ABB RobotStudio station: Pallet_Project_valla_practica.rspag

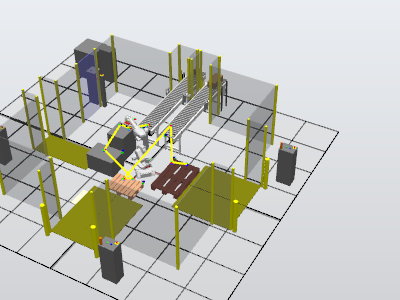
--- station ---
Station Pallet_Project (saved by RobotStudio 24.4.11080.0)
Controller Controler
  mechanical unit ROB_1: IRB1600_10_145__02, 6 joints, base frame (0, 0, 0) mm, rotated rx 0 ry 0 rz 135 deg
Layout (positions relative to the parent item):
  - IRB1600_10_145__02 [mechanism, from %ABB.RobotStudio.Models.IRB1600%\IRB1600_10_145_G_02.rslib] at (0, 0, 0) mm, rotated rx 0 ry 0 rz 135 deg; joint values [0.3434, -0.1552, -0.118, 0, 1.844, -0.442] (rad or m)
  - Half EPAL [part] at (-400, -600, 0) mm, rotated rx 0 ry 0 rz -90 deg, size 600 x 800 x 144 mm
  - ConveyorBox1 [part, from %ABB.RobotStudio.Models.Conveyors%\Conveyor Guide 400.rslib] at (150, 3660, 0) mm, rotated rx 0 ry 0 rz -90 deg
  - ConveyorBox2 [part, from %ABB.RobotStudio.Models.Conveyors%\Conveyor Guide 400.rslib] at (-550, 3660, 0) mm, rotated rx 0 ry 0 rz -90 deg
  - PalletizingVacuumTool [mechanism] at (-560, 265, 1275) mm, rotated rx 180 ry 0 rz 0 deg
      TCP toolVacuum at (0, 0, 175) mm
      links: PalletizingVacuumTool
  - Box1 [part] at (338.5, 3410, 868) mm, size 249 x 499 x 200 mm
  - Box2 [part] at (-353.5, 3575, 868) mm, size 129 x 129 x 200 mm
  - EuroPallet [part, from Components\EuroPalletWood.rslib] at (1400, -600, 0) mm, rotated rx 0 ry 0 rz 90 deg
  - StackingTable [part], size 500 x 600 x 770 mm
  - LinerStand [part], size 800 x 540 x 500 mm
  - SC_Conveyor1 [smart component]
      signals: DO BoxArrived, DI EuroPalletReplaced, DO EuroPalletReplacedOut, DI EuroPalletFull
      connections:
        Source.Executed -> Queue.Enqueue
        PlaneSensor.SensorOut -> Queue.Dequeue
        PlaneSensor.SensorOut -> SC_Conveyor1.BoxArrived
        PlaneSensor.SensorOut -> LogicGate_2.InputA
        LogicGate_2.Output -> Queue_EuroPallet.Enqueue
        LogicGate_2.Output -> Source.Execute
        SimulationEvents.SimulationStarted -> Source.Execute
        SC_Conveyor1.EuroPalletReplaced -> LogicGate_4.InputA
        SC_Conveyor1.EuroPalletFull -> LogicGate_4.InputB
        LogicGate_4.Output -> Queue_EuroPallet.DeleteAll
        LogicGate_4.Output -> SC_Conveyor1.EuroPalletReplacedOut
        Source.Copy => Queue.Back
        Source.Copy => Queue_EuroPallet.Back
    - Source [smart component, from Components\Source.rslib]
        properties: Source=Box1; Copy=(none); Parent=(none); Position=[0.3385 3.39 0.868]; Orientation=[0 0 0]; Transient=true; PhysicsBehavior=-1
    - Queue [smart component, from Components\Queue.rslib]
        properties: Back=(none); Front=(none); Queue={e44fd220-027a-471e-9bb3-a121b85bf4f4};{ee89139f-02ff-44ed-9ba1-277313a75013};{18dc721d-160d-4138-ae65-9469c6fd54a3};{8a7c9217-9ec1-4f6b-adb2-90e3a400ce08};{00ac1772-6055-444c-babb-fd014df5a64d};{22d9b99e-02f4-42e2-875d-e7a2e7a407a6};{801c1d70-c872-49cf-9333-ae7f090aa808};{70a3d2ac-7d8e-4e25-ad4d-efa1d0715e14};{3d190289-ddf5-4821-aefa-1399e7a245df};{fd209546-ad15-4917-a822-45590f893235};{336d7e34-4da5-4704-8767-4e7065a2785d};{a26fb9d1-bd3f-44a5-b61e-f217acd5645d};{35f192af-f0b1-4fcb-92d4-6c5266967521};{7901bdf8-4259-4a58-9fb5-5cf3c990d920};{342c242d-4c7b-4a99-80ec-4606a83008e6};{ba259da1-5c68-49c6-a6dd-ca9a29fb7a6a}; NumberOfObjects=0
    - LinearMover [smart component, from Components\LinearMover.rslib]
        properties: Object=Queue; Direction=[0 -0.001 0]; Speed=0.25; Reference=Global; ReferenceObject=(none)
    - PlaneSensor [smart component, from Components\PlaneSensor.rslib]
        properties: Origin=[0.1885 0.675 0.788]; Axis1=[0.3 0 0]; Axis2=[0 0 0.01]; Tag=(none); SenseMultiple=false; SensedPart=(none)
      - _sensorPart_ [part], size 300 x 0 x 10 mm
    - LogicGate_2 [smart component, from Components\LogicGate.rslib]
        properties: Operator=NOT; Delay=0
    - SimulationEvents [smart component, from Components\SimulationEvents.rslib]
    - Queue_EuroPallet [smart component, from Components\Queue.rslib]
        properties: Back=(none); Front=(none); Queue={ad2057dc-9812-4e01-8eaf-a9764e1c94d2};{23c6148b-879e-4f76-bca6-d4d483c6d4cf};{54fab71e-bcc4-4cca-934a-bbba160b39cc};{b0578ce1-49ea-4c32-a7ca-1e85ec604af9};{947d5054-25d5-43c7-944a-6033d179de93};{94505b46-0998-4fbc-8e5e-e62bbe244ad7};{f8f4ee6a-1769-49de-aeb3-fda26ec8c2f8};{b15d2938-3ac6-4e58-8ecd-de010d23430d};{1b2107f9-d4c6-43db-8eaa-2f076badebbf};{8fdf9589-2ad3-4260-9f23-49ca6aa9f936};{e6f3ceb5-7ecf-422f-9b07-fa91f87616c7};{f8c0f3b0-c392-4387-85be-b0b3c79b7ed2};{b39ef0a3-239a-4eec-87db-20edab27732a};{5504cbc0-0a84-43c9-a60a-8c085a41512d};{4d3e807d-0d48-4360-91da-1f89d28d46d8};{a29bebad-6711-442d-b78a-1822bba72e52};{67d8694a-6ead-419a-ae85-289693a6d2b4};{fe453467-8abc-48a3-b851-8c12c1d7de9d};{6a3e15a0-208f-443f-b6ba-a36fe2c16062};{20e970d1-663c-443e-a64d-d4e9619459f6};{5c8b92e3-60f3-4981-96e7-ca10cb27a842};{db639feb-fd6e-461a-932d-f627d06db2d4};{94b1b66a-00eb-48e1-8857-3db09adf90dc};{618ef0e4-4d6b-4c69-b61e-0bdaa313040e};{043080b5-4091-48b4-bcaf-45ad99666a15};{29caf58f-62f3-4756-8934-f4cc9122e7eb};{7885f061-03ec-4f1c-9005-bd87fa17bd26};{e44fd220-027a-471e-9bb3-a121b85bf4f4};{ee89139f-02ff-44ed-9ba1-277313a75013};{8a7c9217-9ec1-4f6b-adb2-90e3a400ce08};{00ac1772-6055-444c-babb-fd014df5a64d};{22d9b99e-02f4-42e2-875d-e7a2e7a407a6};{801c1d70-c872-49cf-9333-ae7f090aa808};{70a3d2ac-7d8e-4e25-ad4d-efa1d0715e14};{3d190289-ddf5-4821-aefa-1399e7a245df};{fd209546-ad15-4917-a822-45590f893235};{336d7e34-4da5-4704-8767-4e7065a2785d};{a26fb9d1-bd3f-44a5-b61e-f217acd5645d};{35f192af-f0b1-4fcb-92d4-6c5266967521};{7901bdf8-4259-4a58-9fb5-5cf3c990d920};{342c242d-4c7b-4a99-80ec-4606a83008e6}; NumberOfObjects=12
    - LogicGate_4 [smart component, from Components\LogicGate.rslib]
        properties: Operator=AND; Delay=0
  - SC_Gripper [smart component]
      signals: DI Grip
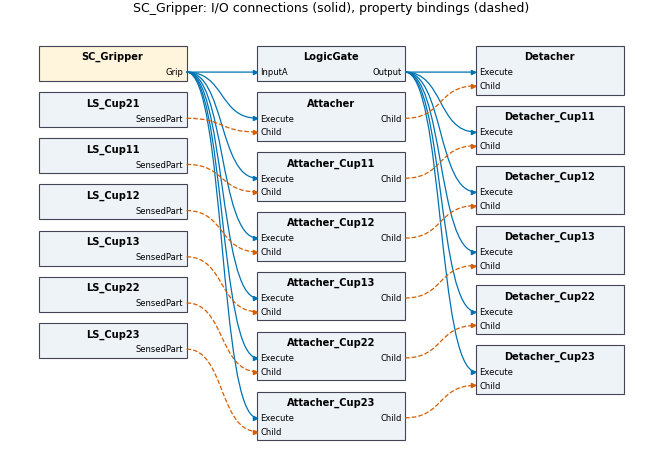
      connections:
        SC_Gripper.Grip -> Attacher.Execute
        SC_Gripper.Grip -> LogicGate.InputA
        LogicGate.Output -> Detacher.Execute
        SC_Gripper.Grip -> Attacher_Cup11.Execute
        LogicGate.Output -> Detacher_Cup11.Execute
        SC_Gripper.Grip -> Attacher_Cup12.Execute
        LogicGate.Output -> Detacher_Cup12.Execute
        SC_Gripper.Grip -> Attacher_Cup13.Execute
        LogicGate.Output -> Detacher_Cup13.Execute
        SC_Gripper.Grip -> Attacher_Cup22.Execute
        LogicGate.Output -> Detacher_Cup22.Execute
        SC_Gripper.Grip -> Attacher_Cup23.Execute
        LogicGate.Output -> Detacher_Cup23.Execute
        LS_Cup21.SensedPart => Attacher.Child
        Attacher.Child => Detacher.Child
        LS_Cup11.SensedPart => Attacher_Cup11.Child
        Attacher_Cup11.Child => Detacher_Cup11.Child
        LS_Cup12.SensedPart => Attacher_Cup12.Child
        Attacher_Cup12.Child => Detacher_Cup12.Child
        LS_Cup13.SensedPart => Attacher_Cup13.Child
        Attacher_Cup13.Child => Detacher_Cup13.Child
        LS_Cup22.SensedPart => Attacher_Cup22.Child
        Attacher_Cup22.Child => Detacher_Cup22.Child
        LS_Cup23.SensedPart => Attacher_Cup23.Child
        Attacher_Cup23.Child => Detacher_Cup23.Child
    - LS_Cup21 [smart component, from Components\LineSensor.rslib] at (190, 265, 153.5) mm, rotated rx 0 ry 0 rz 45 deg
        properties: Start=[-0.597509982704304 0.689429996191639 0.956499992313755]; End=[-0.597509981617333 0.689429995104668 0.924499992313755]; Length=0.032; Radius=0.00331491712707182; Tag=(none); SenseMultiple=false; SensedPart=(none); SensedPoint=[0 0 0]
      - _sensorPart_ [part], size 6.4 x 6.4 x 32 mm
    - Attacher [smart component, from Components\Attacher.rslib]
        properties: Parent=PalletizingVacuumTool; Flange=0; Child=(none); Mount=false; Offset=[0 0 0]; Orientation=[0 0 0]
    - Detacher [smart component, from Components\Detacher.rslib]
        properties: Child=(none); KeepPosition=true
    - LogicGate [smart component, from Components\LogicGate.rslib]
        properties: Operator=NOT; Delay=0
    - LS_Cup11 [smart component, from Components\LineSensor.rslib] at (190, 265, 153.5) mm, rotated rx 0 ry 0 rz 45 deg
        properties: Start=[-0.68943 0.59751 0.9565]; End=[-0.68943 0.59751 0.9245]; Length=0.032; Radius=0.00331; Tag=(none); SenseMultiple=false; SensedPart=(none); SensedPoint=[0 0 0]
      - _sensorPart_ [part], size 6.6 x 6.6 x 32 mm
    - LS_Cup12 [smart component, from Components\LineSensor.rslib] at (190, 265, 153.5) mm, rotated rx 0 ry 0 rz 45 deg
        properties: Start=[-0.57629 0.48437 0.9565]; End=[-0.57629 0.48437 0.9245]; Length=0.032; Radius=0.00331; Tag=(none); SenseMultiple=false; SensedPart=(none); SensedPoint=[0 0 0]
      - _sensorPart_ [part], size 6.6 x 6.6 x 32 mm
    - LS_Cup13 [smart component, from Components\LineSensor.rslib] at (190, 265, 153.5) mm, rotated rx 0 ry 0 rz 45 deg
        properties: Start=[-0.46315 0.37123 0.9565]; End=[-0.46315 0.37123 0.9245]; Length=0.032; Radius=0.00331; Tag=(none); SenseMultiple=false; SensedPart=(none); SensedPoint=[0 0 0]
      - _sensorPart_ [part], size 6.6 x 6.6 x 32 mm
    - LS_Cup22 [smart component, from Components\LineSensor.rslib] at (190, 265, 153.5) mm, rotated rx 0 ry 0 rz 45 deg
        properties: Start=[-0.48437 0.57629 0.9565]; End=[-0.48437 0.57629 0.9245]; Length=0.032; Radius=0.00331; Tag=(none); SenseMultiple=false; SensedPart=(none); SensedPoint=[0 0 0]
      - _sensorPart_ [part], size 6.6 x 6.6 x 32 mm
    - LS_Cup23 [smart component, from Components\LineSensor.rslib] at (190, 265, 153.5) mm, rotated rx 0 ry 0 rz 45 deg
        properties: Start=[-0.37123 0.46315 0.9565]; End=[-0.37123 0.46315 0.9245]; Length=0.032; Radius=0.00331; Tag=(none); SenseMultiple=false; SensedPart=(none); SensedPoint=[0 0 0]
      - _sensorPart_ [part], size 6.6 x 6.6 x 32 mm
    - Attacher_Cup11 [smart component, from Components\Attacher.rslib]
        properties: Parent=PalletizingVacuumTool; Flange=0; Child=(none); Mount=false; Offset=[0 0 0]; Orientation=[0 0 0]
    - Detacher_Cup11 [smart component, from Components\Detacher.rslib]
        properties: Child=(none); KeepPosition=true
    - Attacher_Cup12 [smart component, from Components\Attacher.rslib]
        properties: Parent=PalletizingVacuumTool; Flange=0; Child=(none); Mount=false; Offset=[0 0 0]; Orientation=[0 0 0]
    - Detacher_Cup12 [smart component, from Components\Detacher.rslib]
        properties: Child=(none); KeepPosition=true
    - Attacher_Cup13 [smart component, from Components\Attacher.rslib]
        properties: Parent=PalletizingVacuumTool; Flange=0; Child=(none); Mount=false; Offset=[0 0 0]; Orientation=[0 0 0]
    - Detacher_Cup13 [smart component, from Components\Detacher.rslib]
        properties: Child=(none); KeepPosition=true
    - Attacher_Cup22 [smart component, from Components\Attacher.rslib]
        properties: Parent=PalletizingVacuumTool; Flange=0; Child=(none); Mount=false; Offset=[0 0 0]; Orientation=[0 0 0]
    - Detacher_Cup22 [smart component, from Components\Detacher.rslib]
        properties: Child=(none); KeepPosition=true
    - Attacher_Cup23 [smart component, from Components\Attacher.rslib]
        properties: Parent=PalletizingVacuumTool; Flange=0; Child=(none); Mount=false; Offset=[0 0 0]; Orientation=[0 0 0]
    - Detacher_Cup23 [smart component, from Components\Detacher.rslib]
        properties: Child=(none); KeepPosition=true
  - SC_Conveyor2 [smart component]
      signals: DO BoxArrived, DI HalfPalletReplaced, DI HalfPalletFull, DO HalfPalletReplacedOut
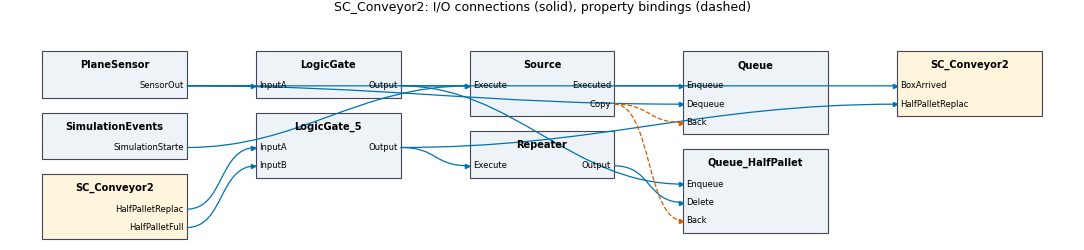
      connections:
        Source.Executed -> Queue.Enqueue
        PlaneSensor.SensorOut -> Queue.Dequeue
        PlaneSensor.SensorOut -> SC_Conveyor2.BoxArrived
        PlaneSensor.SensorOut -> LogicGate.InputA
        SimulationEvents.SimulationStarted -> Source.Execute
        LogicGate.Output -> Queue_HalfPallet.Enqueue
        LogicGate.Output -> Source.Execute
        Repeater.Output -> Queue_HalfPallet.Delete
        SC_Conveyor2.HalfPalletReplaced -> LogicGate_5.InputA
        SC_Conveyor2.HalfPalletFull -> LogicGate_5.InputB
        LogicGate_5.Output -> Repeater.Execute
        LogicGate_5.Output -> SC_Conveyor2.HalfPalletReplacedOut
        Source.Copy => Queue.Back
        Source.Copy => Queue_HalfPallet.Back
    - Source [smart component, from Components\Source.rslib]
        properties: Source=Box2; Copy=(none); Parent=(none); Position=[-0.3535 3.575 0.868]; Orientation=[0 0 0]; Transient=true; PhysicsBehavior=-1
    - Queue [smart component, from Components\Queue.rslib]
        properties: Back=(none); Front=(none); Queue={d41f34b8-4a20-475c-95ba-460bc2504caf};{5a16ad96-9ff6-44fe-ab59-6bd35466d4d1};{0f18d6dc-c4e6-4c44-9757-559d16fce4ae};{b2c7b4bf-0d60-42df-8ee4-abc0a1068e12};{8d30a67c-a063-4d22-a747-3e9a99cdef41};{1409c1e2-dbf3-49bd-b776-9bd8588f9165};{e3acce53-8455-4384-b1ac-df89878ccd5c};{87db3190-4758-4831-8d2c-d9fdcd68b36e};{469258bd-729a-49fe-bc80-31f695b1b400};{4c1b5bae-9eaf-40c3-874b-2538b6841d7a};{46ba244e-445c-470d-b6ca-5e376dcf2b7e};{e5ec3e26-f6d7-4e6f-b347-541b5d6ec99e}; NumberOfObjects=0
    - LinearMover [smart component, from Components\LinearMover.rslib]
        properties: Object=Queue; Direction=[0 -0.001 0]; Speed=0.25; Reference=Global; ReferenceObject=(none)
    - PlaneSensor [smart component, from Components\PlaneSensor.rslib]
        properties: Origin=[-0.5035 0.675 0.788]; Axis1=[0.3 0 0]; Axis2=[0 0 0.01]; Tag=(none); SenseMultiple=false; SensedPart=(none)
      - _sensorPart_ [part], size 300 x 0 x 10 mm
    - LogicGate [smart component, from Components\LogicGate.rslib]
        properties: Operator=NOT; Delay=0
    - SimulationEvents [smart component, from Components\SimulationEvents.rslib]
    - Queue_HalfPallet [smart component, from Components\Queue.rslib]
        properties: Back=(none); Front=(none); Queue={f5edb1ce-3bf5-426a-a389-0b0047efa949};{5ce0816a-b692-43c6-82f7-492eb3fc1c7c};{ad3ef4b5-2c59-4daa-9658-0c77e5efb67d};{c9c476d0-74ff-4b18-bfb3-2d6c852b8493};{1bf865c6-1649-4319-b5ff-cd81faaa6069};{f626778c-15a6-4059-b27a-7c8f9da4f34f};{a60dd0dd-490e-48fe-bb32-16f415136b44};{4ec9b3b2-e4a8-4d14-aea0-9552a35d2afd};{38bc6a68-8d9e-44a7-a5f0-badb214ea710};{f9543542-377a-43f1-9613-018dced76680};{486b4c2f-b225-4486-b430-5ab7d813c599};{7da52d9e-9053-4b1a-839c-0aedc5495cc7};{c2400356-fde5-4523-9dc7-d26788098951};{75099568-1fe6-4c34-8328-63fd42144c3b};{8ca6c374-2d39-4938-8324-38c48ae4f51d};{f3c160ab-6f5f-460b-8b54-c2c3b0bc175f};{1c289510-9a29-4e1c-b603-54b7a0027260};{d39da69b-e59a-4ace-85a5-bba54583b01c};{bc328c62-4bf3-4a57-965c-0c93e0ee296d};{60f4dcb3-d366-4d0b-b05a-5b2073fcd9e8};{44334a49-cf52-4d95-9964-3bb568ce732d};{f9240695-1965-47e5-bcd4-644ec5904899};{72a970fd-f238-4ac5-b811-00686975bc20};{bd297b2a-4ad7-44fa-87c8-1ac40b0d2fbf};{3dafa88d-62b0-429f-9c75-c8c7bde09fc6};{a7d8f176-4e9d-4819-8805-982bee0c310d};{72ae6bb6-3373-4f60-a321-dfdc0981c562};{fff16105-3d56-4b21-a888-399904fd95d4};{56e4abf9-acd4-4a00-b067-52a58200d221};{2eb8ae55-b553-4f83-b65d-07c27c701dd6};{dfb05241-1220-45e8-b584-1559777c0125};{49a2c23a-27ea-4b0b-af5c-f9d01014f642};{0adfb5d7-4fd0-41be-8361-c42c9d28ca51};{8cf74624-f46b-49ca-a524-038ddb88ba0f};{bde2cdc4-b3e4-48fe-8333-d64185b5a8e7};{d17564c2-89d4-4b4f-8596-5dca9165a286};{6fec26e7-cb1b-4d74-b4a6-8ed7a2eb81a6};{e04d8697-cc19-4df5-b7fa-dff41516820c};{134714af-70a5-49a3-8b99-ea847d1ef329};{23aa8eff-aaeb-4079-b6e6-9fe5f0b7799c};{0091a76d-e23e-4382-9bf3-a427b049953f};{fdc2abc9-40b2-462e-8472-b1d156765a68};{8dc86a38-8dcf-454b-a79a-3f5e6d46a581};{f9226736-fe9f-4ce5-82b5-97fc8f487c87};{8d0584df-2d5d-4d5a-bd5b-c865cb85c145};{fef2818e-b6b9-47fe-bf8a-83543bb000b1};{5ac98beb-c6da-4ea7-80b2-93f7dacce3e5};{443aad51-6408-442e-915b-2ecfdc577e14};{51b93794-f199-43f0-a14e-6aec3c171668};{885be8a6-b854-423c-907a-f456456dba07};{dcbbb2a9-79f1-4094-9b60-3ac8a0070454};{86281ae9-2d9e-4987-a35e-6d6a445e8875};{9f234810-50d8-438d-8980-298a5844ac16};{4c457525-5ea0-4a08-bfa0-e2a51e8a57a9};{d60c358c-9baa-495a-a755-dc91e6e5630d};{cba8d61a-9576-424b-b333-8920ed1679e6};{fffcb6aa-6454-497e-a713-529b874f7300};{8c292b69-8603-4861-ab75-8c5041fc1228};{be74d22e-2a24-4d51-b9be-30cb4581f5e4};{9c8c849d-9d7a-4314-9edc-0c9679818308};{51cbe104-3a08-4083-a326-34fc650c90a2};{8d9adc3a-e0d0-484f-8727-84b992719000};{9a2b47ee-5540-43de-9a30-89f96a258b35};{cfb929ec-bf51-45d3-8071-aea9b14bf075};{867175b9-70b9-45ce-970c-131187ba34ca};{173082af-f5ae-4239-8a69-7ad684951e00};{b2c9da23-dceb-4407-8f95-0d503246dac3};{f0464754-db31-42ef-9c41-8ce46a4a0971};{6b29df5c-760d-4911-84dd-92d25b30bb71};{8cf0ae3d-fbb1-4655-8db9-abf8850d857b};{fcdbf145-8b27-4e5e-9241-3719648eab1d};{78faf9d5-81df-4a41-87f3-b1a514ef17c7};{3a4d91ff-54a0-485c-9c99-c5554510e37a};{c01a110e-561d-45dd-b1c3-10d79a4111a8};{63ad2c6d-e580-44e3-9dfc-7106564b7944};{ccc00ef2-4c06-4459-824e-6f17fc3bacb7};{b81e233c-b00c-4cd7-b93a-2cecac8f8dc1};{398e0c88-f727-4b42-8f39-aaa6835500b7};{fc631786-067a-487d-abac-51fcb0c6dd41};{cf6ca633-09f3-4f3b-9435-b43791280bff};{74bed72d-6a54-4305-87bd-9ad3015ece89};{bb2cc45e-a4eb-4ab2-9ef7-f371e7fbe706};{dd82f376-2e09-4208-84ad-5816bed92574};{e392904e-f13d-4939-a056-7304ff0c878c};{3e44c1eb-892b-48b7-9eef-a2eb6a338ec4};{67a95a53-b6c9-4e7f-9fd4-7782a33b0ce9};{b907a4a1-1349-44c4-99ca-3ea2b14844a2};{27bb147c-485e-4ba4-8918-f2e2468aa20b};{4158548c-0e01-4059-887d-ce75515d9624};{bdcc830f-a4a4-4608-9c6a-3968c3b56955};{8ac99da1-daa1-4239-8c24-2cbcd0fbbccf};{eceb8029-a656-40f5-a7a3-28283ded6e47};{06ec9c8e-bd56-4499-906c-965bdc743b38};{bc8629f4-be69-483d-a42b-bd5694970e3a};{91c33ad6-79d6-4ff7-b807-aaf3d283071a};{bbff1efe-9f6d-4f6e-9e11-7159709d58b9};{d8345c1f-8548-4957-9dd2-2c7a65aadcb5};{297050bf-6bdd-4149-9774-639d35df4273};{9047bf3c-f537-46c2-88b1-9fd2d5954a0b};{5951cc55-a535-4f63-8005-57734053514f};{4bb3aaf8-1744-440d-8239-fce36f67cc2c};{eb7c6c5d-8b86-4d0e-b965-01e8cc90c395};{da949c7c-7130-455a-a5de-886672c52ec3};{04b934b1-2ca6-4947-808f-8dc968a55eb4};{d4940027-1ade-4406-ae0f-2cc92eccc776};{37dc3e2f-17e0-406e-80b6-d473aa1734f3};{09cf0d3f-945d-4baa-a296-e9bd267df3af};{8a94d3e3-b0e3-42c4-90bd-ba639180af74};{049eaf7e-723f-484a-b080-48153e5693e0};{2c2227db-366e-4824-818a-8891fec9d39b};{78a4912a-e493-4427-95eb-ed4a7e141f53};{8b1769a4-052b-4f7f-be48-9c2315e00515};{4bb9eccd-54a8-444b-8b85-f69dc35199f7};{5d771788-ec0f-48bc-9cbe-993fb932c8ea};{021fadd8-996c-49c9-9ff6-8a460f8c358b};{e61d541c-af94-4f27-b95d-aac3b95a1cd9};{a0819d77-e800-4559-87f4-c656405fa595};{003f191f-efb3-43bb-b7aa-33133ee6defd};{3abac3eb-5c5c-4177-b0e4-5f71daa2fcd7};{f4938c82-19bc-4592-9d12-63feb2c87ac4};{2b776e4a-67ea-499c-995e-bce8af0160a7};{c9a77fd9-e2d1-4dbf-8d0e-8377c4665448};{62bb8355-d295-4471-b563-b6f46f05c8b1};{55201944-7d05-43e8-bd24-433bd506e7b6};{76821f68-2096-4060-b9d6-b9517b2f6dc5};{e09ad2c9-6668-417d-a6ce-db14256207b6};{ca102da5-219d-413a-ab81-6e9821c26e06};{c588302c-8cce-44a8-91f3-143c0654eb27};{2202393d-e22d-4f8c-8a1d-1cc72ba5cca5};{be80ae30-a6c8-4766-bc6b-bfe80846e161};{25475f3f-ef68-45ff-aa3c-0ea04c10e4e7};{498aca50-8032-4c24-8147-7ec56c07f7a0};{b4a07b3f-831d-4f53-9343-c16642fe3bc1};{8bd52ab4-c09d-4b2d-8603-56cbb3c77529};{6f1069cf-970f-4855-ba49-8ae785987118};{b667b62f-e5f1-478a-9bad-dc3725da1d04};{86e8e265-466a-4a6e-8b5e-b128819dda1c};{4df69d20-688f-43ef-bee0-112974bed187};{182f9b53-f0c9-4414-a7de-97eac4ce486a};{514b0f5e-2197-4430-9c07-cfb19e0d92ad};{359ebd0e-6711-4070-a5d3-939e22007801};{d67847b8-c0ad-4246-ba67-b0d24865206c};{197fb8bb-a523-4e0e-8be7-47cc1723a988};{142dd6b6-47a3-4a32-99f8-9706d11eb229};{1a8963b6-e72b-4e55-95a7-15d5212af876};{42897a06-6f96-425a-a387-4cefe2eac35b};{d78e4ef6-3fce-473d-bfe7-e529abd3d695};{e0b062dd-5846-40f4-b32c-2a1ab6da1894};{4c4aa1cf-e61f-45c1-9c13-55311062428a};{a0d6a9a4-70e0-4c3a-ae7d-eaf5e5bb2112};{bc16083c-a858-482a-a879-7c8861b2473f};{64ab26ad-0b46-4ced-ab7f-1cfee37682ad};{2165d0dd-c254-4ebf-83cc-be68d523d748};{44491ebe-5cdd-46fe-a821-5ec7c79b16a0};{ddfa3b39-85f7-4855-9203-7f7a6cdd8093};{137fe74d-152f-4b74-9f93-d403c4354bb3};{82ca252e-23ba-4001-8e89-7b23c4c78f2e};{062cf830-d27c-401d-a518-3a9fb83d9537};{610befe8-cd72-44d2-af6b-444eaea3df38};{cf0b5eb3-bda2-46b1-b486-9a887917bee5};{a53ebe9a-d0a3-4afd-b901-97852e5709fd};{8b5126a5-3700-41cc-bd9b-a335d093d62b};{1a031046-3bf3-47b0-bf1d-63f834d0f0bf};{32ae9498-3575-4e70-954e-9800b2c7ed18};{ee3cbed5-90f6-47a6-8d41-8a31a6a9b52f};{f52f3a91-5bd6-47b6-a1f8-92ea9cad0f19};{b2f50ce9-01bf-4326-9e7f-81a685c29d51};{db908664-ce90-4d8d-99e6-8cad1d25b072};{ce174d6d-3e8c-4abc-807c-2e034a05442b};{6b3f855e-a78e-40d1-a8e8-dc264647088d};{cde41289-1748-48b7-acac-ba93367ef0bd};{23d0bcac-3df5-4d02-9989-7a0bd57a2c5a};{7d6ef79f-31a3-4faa-a3c8-24190ad66021};{148a4a69-c3f4-4709-9c4e-248710d37209};{3a43107f-6ec5-42b1-bdab-65f53844f08b};{688ca237-9237-4c0d-9f6a-943bdaf2a54e};{b0c649b2-1e95-4926-b3f4-7de3359bf184};{775c86bc-3b84-4fb2-a4b9-0c2b4654e980};{d13aeccf-57c6-48c5-8ccb-e0d83af0bf52};{b23f60bf-e49d-4af6-aa11-454509134c6f};{0a5e5d93-42f5-44d1-80bb-87a9dcd65f82};{03917fb8-4550-48ea-aade-cad2296182d4};{69fc404e-23e5-4586-8106-722a8d502888};{efd93624-9dc8-470c-9ca5-761da3b13f64};{3161c526-c456-4198-a8e9-6ba9dc97d08d};{1f8ccdfc-77be-4eb2-b50b-b6f397d92aac};{cb468d26-4eaa-493f-84ab-65bfcf757383};{bd96b98c-b60d-47b5-9e29-6a1dfadd5ba3};{35cfaa90-f083-49e1-b726-d654efc82f59};{60633137-d3a6-410f-a68f-c3960af01eec};{b8faed0a-d8df-4dd7-a7c6-c20d690a082c};{469fa596-a3ad-4a84-8b8e-6f04cb45c4e6};{543f5b18-19fb-410f-92c3-c1199be26dff};{1f728d5f-b843-4df0-b352-629d14987f1c};{12323632-ef84-4060-aa52-b2f1987c73f3};{062735fc-4a51-4d85-95c2-a683477f8e45};{444b3eac-f57f-4356-8db0-63ce6624c93d};{325a86c2-b1da-40af-a81a-eb00a2886e08};{73c79afd-8798-467b-80dd-9e32e888d88c};{f243e6a9-0264-46d4-8a6c-a8c2b4c42193};{f7d0602e-30eb-44b6-b654-6cdc5756be59};{ad2ed4ca-30e0-4614-a0d8-f4fea7ef6fce};{bab6a964-a4d0-4eed-9c33-fa686721e8e3};{fb67aacc-6733-43ed-a4db-7a6425d2d60c};{6421a31f-3a82-4b20-9081-df48bb7907b5};{8ff8c115-8e7b-4406-a53a-edf3873335b8};{5ac3eee3-ab48-4a86-8294-3ac57f94e03f};{d41f34b8-4a20-475c-95ba-460bc2504caf};{5a16ad96-9ff6-44fe-ab59-6bd35466d4d1};{0f18d6dc-c4e6-4c44-9757-559d16fce4ae};{b2c7b4bf-0d60-42df-8ee4-abc0a1068e12};{8d30a67c-a063-4d22-a747-3e9a99cdef41};{1409c1e2-dbf3-49bd-b776-9bd8588f9165};{e3acce53-8455-4384-b1ac-df89878ccd5c};{87db3190-4758-4831-8d2c-d9fdcd68b36e};{469258bd-729a-49fe-bc80-31f695b1b400};{4c1b5bae-9eaf-40c3-874b-2538b6841d7a};{46ba244e-445c-470d-b6ca-5e376dcf2b7e}; NumberOfObjects=78
    - Repeater [smart component, from Components\Repeater.rslib]
        properties: Count=72
    - LogicGate_5 [smart component, from Components\LogicGate.rslib]
        properties: Operator=AND; Delay=0
  - Liner_01 [part] at (-900, -2000, 0) mm, size 800 x 540 x 10 mm
  - SC_Liners [smart component]
      signals: DI LinersRefilled, DI LinerStackEmpty, DI PalletReplaced, DO LinersRefilledOut
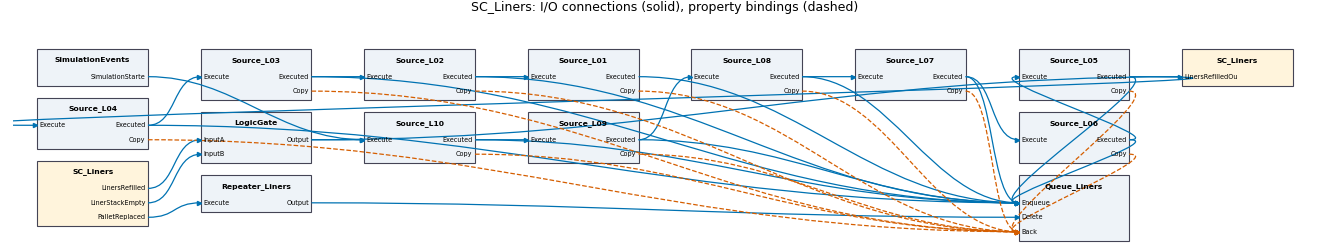
      connections:
        SimulationEvents.SimulationStarted -> Source_L10.Execute
        Source_L10.Executed -> Queue_Liners.Enqueue
        Source_L10.Executed -> Source_L09.Execute
        Source_L09.Executed -> Queue_Liners.Enqueue
        Source_L09.Executed -> Source_L08.Execute
        Source_L08.Executed -> Queue_Liners.Enqueue
        Source_L08.Executed -> Source_L07.Execute
        Source_L07.Executed -> Queue_Liners.Enqueue
        Source_L07.Executed -> Source_L06.Execute
        Source_L06.Executed -> Queue_Liners.Enqueue
        Source_L06.Executed -> Source_L05.Execute
        Source_L05.Executed -> Queue_Liners.Enqueue
        Source_L05.Executed -> Source_L04.Execute
        Source_L04.Executed -> Queue_Liners.Enqueue
        Source_L04.Executed -> Source_L03.Execute
        Source_L03.Executed -> Queue_Liners.Enqueue
        Source_L03.Executed -> Source_L02.Execute
        Source_L02.Executed -> Queue_Liners.Enqueue
        Source_L02.Executed -> Source_L01.Execute
        Source_L01.Executed -> Queue_Liners.Enqueue
        SC_Liners.LinersRefilled -> LogicGate.InputA
        SC_Liners.LinerStackEmpty -> LogicGate.InputB
        LogicGate.Output -> SC_Liners.LinersRefilledOut
        LogicGate.Output -> Source_L10.Execute
        SC_Liners.PalletReplaced -> Repeater_Liners.Execute
        Repeater_Liners.Output -> Queue_Liners.Delete
        Source_L10.Copy => Queue_Liners.Back
        Source_L09.Copy => Queue_Liners.Back
        Source_L08.Copy => Queue_Liners.Back
        Source_L07.Copy => Queue_Liners.Back
        Source_L06.Copy => Queue_Liners.Back
        Source_L05.Copy => Queue_Liners.Back
        Source_L04.Copy => Queue_Liners.Back
        Source_L03.Copy => Queue_Liners.Back
        Source_L02.Copy => Queue_Liners.Back
        Source_L01.Copy => Queue_Liners.Back
    - Source_L10 [smart component, from Components\Source.rslib]
        properties: Source=Liner_01; Copy=(none); Parent=(none); Position=[-1.3 -0.7 0.59]; Orientation=[0 0 0]; Transient=true; PhysicsBehavior=-1
    - Source_L09 [smart component, from Components\Source.rslib]
        properties: Source=Liner_01; Copy=(none); Parent=(none); Position=[-1.3 -0.7 0.58]; Orientation=[0 0 0]; Transient=true; PhysicsBehavior=-1
    - Queue_Liners [smart component, from Components\Queue.rslib]
        properties: Back=(none); Front=(none); Queue={4b76874b-49d8-40e7-b1bf-01d8cc753daf};{f1bc3993-1843-4745-a916-cd233907ef8f};{7d1f5471-804d-47e8-8c82-babb94078c4f};{35f64396-636a-40cf-85a6-257e77a6ae60};{2aedaf41-8ae8-41b0-9db2-9de3ceaf795b};{436fe240-c7f2-42eb-89c0-1cd4aff7e3ff};{e7949e0b-2972-403e-9743-54dc0693f87f};{59bd0fcf-8828-44fb-b45a-84ebd2dc8c3d};{59a7902e-96f8-4e0e-b708-dc1c92c26f66};{1f249118-cd38-42be-b8a7-d3254198917b};{33f64cea-21b7-4476-9a21-b1850c845c4c};{6d880d10-0093-43e7-8014-139534ada452};{8432c400-4781-49f7-aa39-fa2dc6e98a0f};{61e97684-8218-4ac6-a060-0ca69cab5273};{78371439-59e8-482d-8147-9dece47c4b3d};{5351f5ec-037c-4625-be08-d259f2f0dab9};{1728b901-d880-497f-a9dc-fc428da0f52d};{94273ab4-5060-46c3-80b2-362935833b91};{3e6b5fa6-26e1-42c5-aada-9e85978ab4cf};{89a16311-d9f3-4be9-874c-e3d1f0939d0f};{01a3968c-dc38-41a8-821e-9eb7eb9ddcb6};{f6651478-43f4-42ca-bae1-f1f503b6b42a};{2f17a5c0-632c-4a5a-aea8-f6e212c5841b};{69ef7725-acb4-4562-810a-a97a14cbd53c};{704c2d3b-24d3-475f-8d25-b6b26e7fec9c};{f2ed20fd-a82f-4770-a0af-12c07cfbfa73};{d8dcd6ae-656a-4bcc-8399-251caf5a0e2f};{4f1be6df-21fc-4212-9b62-51a6ddf46789};{f83a54dd-86e1-4b51-ad4c-f3092acc29ee};{534771e2-1ace-4b39-b107-fcece75fcd88};{006ab1e9-1667-49eb-a3fc-9daf3d261695};{5cff699e-b7b2-4f06-b0dd-3aa3a2565d54};{62b4127a-2a9b-4d56-a22d-ac07527ab970};{72a0e263-fa92-4955-bee8-75cd8e7bcda3};{2f5c7ce6-cc96-4025-8b6f-42fc8d1c53de};{a007f585-8c80-40f3-9f22-79fa01fd41be};{7214a086-acb6-4dc9-80a5-5db08c6fb4b9};{12bb64d4-b495-4b48-a9c8-db9791f029e3};{32b5cfa5-8504-4b44-a4bf-b1b8b1e80030};{60a53e66-30e6-4fde-a9d2-765474ab08f2};{31019e2a-21cb-4e2c-9cdb-7de64fe533e9};{09e6c226-ece6-4f81-9df3-2592efd7026c}; NumberOfObjects=10
    - SimulationEvents [smart component, from Components\SimulationEvents.rslib]
    - Source_L08 [smart component, from Components\Source.rslib]
        properties: Source=Liner_01; Copy=(none); Parent=(none); Position=[-1.3 -0.7 0.57]; Orientation=[0 0 0]; Transient=true; PhysicsBehavior=-1
    - Source_L07 [smart component, from Components\Source.rslib]
        properties: Source=Liner_01; Copy=(none); Parent=(none); Position=[-1.3 -0.7 0.56]; Orientation=[0 0 0]; Transient=true; PhysicsBehavior=-1
    - Source_L06 [smart component, from Components\Source.rslib]
        properties: Source=Liner_01; Copy=(none); Parent=(none); Position=[-1.3 -0.7 0.55]; Orientation=[0 0 0]; Transient=true; PhysicsBehavior=-1
    - Source_L05 [smart component, from Components\Source.rslib]
        properties: Source=Liner_01; Copy=(none); Parent=(none); Position=[-1.3 -0.7 0.54]; Orientation=[0 0 0]; Transient=true; PhysicsBehavior=-1
    - Source_L04 [smart component, from Components\Source.rslib]
        properties: Source=Liner_01; Copy=(none); Parent=(none); Position=[-1.3 -0.7 0.53]; Orientation=[0 0 0]; Transient=true; PhysicsBehavior=-1
    - Source_L03 [smart component, from Components\Source.rslib]
        properties: Source=Liner_01; Copy=(none); Parent=(none); Position=[-1.3 -0.7 0.52]; Orientation=[0 0 0]; Transient=true; PhysicsBehavior=-1
    - Source_L02 [smart component, from Components\Source.rslib]
        properties: Source=Liner_01; Copy=(none); Parent=(none); Position=[-1.3 -0.7 0.51]; Orientation=[0 0 0]; Transient=true; PhysicsBehavior=-1
    - Source_L01 [smart component, from Components\Source.rslib]
        properties: Source=Liner_01; Copy=(none); Parent=(none); Position=[-1.3 -0.7 0.5]; Orientation=[0 0 0]; Transient=true; PhysicsBehavior=-1
    - LogicGate [smart component, from Components\LogicGate.rslib]
        properties: Operator=AND; Delay=0
    - Repeater_Liners [smart component, from Components\Repeater.rslib]
        properties: Count=2
  - Door_Maintenance [part], size 20 x 800 x 2000 mm
  - LightCurtain_EuroPallet_Emitter [part], size 50 x 50 x 2000 mm
  - LightCurtain_EuroPallet_Receiver [part], size 50 x 50 x 2000 mm
  - LightCurtain_HalfPallet_Emitter [part], size 50 x 50 x 2000 mm
  - LightCurtain_HalfPallet_Receiver [part], size 50 x 50 x 2000 mm
  - LightCurtain_LinerBay_Emitter [part], size 50 x 50 x 2000 mm
  - LightCurtain_LinerBay_Receiver [part], size 50 x 50 x 2000 mm
  - LightCurtain_Conv1_Emitter [part], size 50 x 50 x 450 mm
  - LightCurtain_Conv1_Receiver [part], size 50 x 50 x 450 mm
  - LightCurtain_Conv2_Emitter [part], size 50 x 50 x 450 mm
  - LightCurtain_Conv2_Receiver [part], size 50 x 50 x 450 mm
  - MutingSensor_Conv1_A [part], size 30 x 30 x 900 mm
  - MutingSensor_Conv1_B [part], size 30 x 30 x 900 mm
  - MutingSensor_Conv2_A [part], size 30 x 30 x 900 mm
  - MutingSensor_Conv2_B [part], size 30 x 30 x 900 mm
  - SafetyMat_EuroPallet [part], size 1650 x 1800 x 15 mm
  - SafetyMat_HalfPallet [part], size 1500 x 1850 x 15 mm
  - SafetyMat_LinerBay [part], size 1750 x 740 x 15 mm
  - PalletStop_Euro_1 [part], size 40 x 100 x 80 mm
  - PalletStop_Euro_2 [part], size 40 x 100 x 80 mm
  - PalletStop_Half_1 [part], size 100 x 40 x 80 mm
  - PalletStop_Half_2 [part], size 100 x 40 x 80 mm
  - OperatorStation_EuroPallet [part], size 400 x 300 x 1100 mm
  - OperatorStation_HalfPallet [part], size 400 x 300 x 1100 mm
  - OperatorStation_LinerBay [part], size 400 x 300 x 1100 mm
  - OperatorStation_General [part], size 400 x 300 x 1100 mm
  - OperatorStation_Door [part], size 300 x 300 x 1100 mm
  - EStopPost_Inside [part], size 100 x 100 x 1100 mm
  - IRC5_Cabinet [part], size 725 x 710 x 970 mm
  - DoorSensor_Eden_Actuator [part], size 30 x 40 x 60 mm
  - DoorSensor_Eden_Sensor [part], size 30 x 40 x 60 mm
  - EStopBase_EuroPallet [part], size 80 x 80 x 5 mm
  - EStopBase_HalfPallet [part], size 80 x 80 x 5 mm
  - EStopBase_LinerBay [part], size 80 x 80 x 5 mm
  - EStopBase_General [part], size 80 x 80 x 5 mm
  - EStopBase_Door [part], size 80 x 80 x 5 mm
  - EStopBase_Inside [part], size 80 x 80 x 5 mm
  - Bumper_EuroPallet_1 [part], size 114 x 114 x 1000 mm
  - Bumper_EuroPallet_2 [part], size 114 x 114 x 1000 mm
  - Bumper_HalfPallet_1 [part], size 114 x 114 x 1000 mm
  - Bumper_HalfPallet_2 [part], size 114 x 114 x 1000 mm
  - MutingLamp_Conv1 [part], size 60 x 60 x 100 mm
  - MutingLamp_Conv2 [part], size 60 x 60 x 100 mm
  - Lamp_EuroPalletFull [part], size 60 x 59.8 x 200 mm
  - Lamp_HalfPalletFull [part], size 60 x 59.8 x 200 mm
  - Lamp_LinerStackEmpty [part], size 60 x 59.8 x 200 mm
  - Button_EuroPalletReplaced [part], size 40 x 39.9 x 20 mm
  - Button_HalfPalletReplaced [part], size 40 x 39.9 x 20 mm
  - Button_LinersRefilled [part], size 40 x 39.9 x 20 mm
  - ResetButton_EuroPallet [part], size 40 x 39.9 x 20 mm
  - ResetButton_HalfPallet [part], size 40 x 39.9 x 20 mm
  - ResetButton_LinerBay [part], size 40 x 39.9 x 20 mm
  - ResetButton_Door [part], size 40 x 39.9 x 20 mm
  - EStop_EuroPallet [part], size 40 x 40 x 30 mm
  - EStop_HalfPallet [part], size 40 x 40 x 30 mm
  - EStop_LinerBay [part], size 40 x 40 x 30 mm
  - EStop_General [part], size 40 x 40 x 30 mm
  - EStop_Door [part], size 40 x 40 x 30 mm
  - EStop_Inside [part], size 40 x 40 x 30 mm
  - Safety_Fence [graphiccomponentgroup]
    - Fence_Corridor_Euro_1 [part], size 500 x 20 x 2000 mm
    - Fence_Corridor_Euro_2 [part], size 500 x 20 x 2000 mm
    - Fence_Corridor_Half_1 [part], size 20 x 500 x 2000 mm
    - Fence_Corridor_Half_2 [part], size 20 x 500 x 2000 mm
    - Fence_Corridor_Liner_1 [part], size 500 x 20 x 2000 mm
    - Fence_Corridor_Liner_2 [part], size 500 x 20 x 2000 mm
    - Fence_Panel_E1 [part], size 20 x 1650 x 2000 mm
    - Fence_Panel_E2 [part], size 20 x 1650 x 2000 mm
    - Fence_Panel_N1 [part], size 1931.5 x 20 x 2000 mm
    - Fence_Panel_N2 [part], size 162 x 20 x 2000 mm
    - Fence_Panel_N3 [part], size 1946.5 x 20 x 2000 mm
    - Fence_Panel_S1 [part], size 1800 x 20 x 2000 mm
    - Fence_Panel_S2 [part], size 1800 x 20 x 2000 mm
    - Fence_Panel_W1 [part], size 20 x 1750 x 2000 mm
    - Fence_Panel_W2 [part], size 20 x 960 x 2000 mm
    - Fence_Panel_W3 [part], size 20 x 850 x 2000 mm
    - Fence_Post_01 [part], size 60 x 60 x 2000 mm
    - Fence_Post_02 [part], size 60 x 60 x 2000 mm
    - Fence_Post_03 [part], size 60 x 60 x 2000 mm
    - Fence_Post_04 [part], size 60 x 60 x 2000 mm
    - Fence_Post_05 [part], size 60 x 60 x 2000 mm
    - Fence_Post_06 [part], size 60 x 60 x 2000 mm
    - Fence_Post_07 [part], size 60 x 60 x 2000 mm
    - Fence_Post_08 [part], size 60 x 60 x 2000 mm
    - Fence_Post_09 [part], size 60 x 60 x 2000 mm
    - Fence_Post_10 [part], size 60 x 60 x 2000 mm
    - Fence_Post_11 [part], size 60 x 60 x 2000 mm
    - Fence_Post_12 [part], size 60 x 60 x 2000 mm
    - Fence_Post_13 [part], size 60 x 60 x 2000 mm
    - Fence_Post_14 [part], size 60 x 60 x 2000 mm
    - Fence_Post_15 [part], size 60 x 60 x 2000 mm
    - Fence_Post_16 [part], size 60 x 60 x 2000 mm
    - Fence_Post_17 [part], size 60 x 60 x 2000 mm
    - Fence_Post_18 [part], size 60 x 60 x 2000 mm
    - Fence_Post_19 [part], size 60 x 60 x 2000 mm
    - Fence_Post_20 [part], size 60 x 60 x 2000 mm
    - Fence_Tunnel_Conv1_1 [part], size 20 x 500 x 2000 mm
    - Fence_Tunnel_Conv1_2 [part], size 20 x 500 x 2000 mm
    - Fence_Tunnel_Conv1_Low [part], size 530 x 20 x 700 mm
    - Fence_Tunnel_Conv1_Top [part], size 530 x 20 x 980 mm
    - Fence_Tunnel_Conv2_1 [part], size 20 x 500 x 2000 mm
    - Fence_Tunnel_Conv2_2 [part], size 20 x 500 x 2000 mm
    - Fence_Tunnel_Conv2_Low [part], size 530 x 20 x 700 mm
    - Fence_Tunnel_Conv2_Top [part], size 530 x 20 x 980 mm
Attachment: PalletizingVacuumTool is attached to IRB1600_10_145__02 / Link6
Attachment: LS_Cup21 is attached to PalletizingVacuumTool / PalletizingVacuumTool
Attachment: LS_Cup12 is attached to PalletizingVacuumTool / PalletizingVacuumTool
Attachment: LS_Cup13 is attached to PalletizingVacuumTool / PalletizingVacuumTool
Attachment: LS_Cup22 is attached to PalletizingVacuumTool / PalletizingVacuumTool
Attachment: LS_Cup23 is attached to PalletizingVacuumTool / PalletizingVacuumTool
Attachment: LS_Cup11 is attached to PalletizingVacuumTool / PalletizingVacuumTool
Collision set Conjunto de colisión_1: IRB1600_10_145__02, PalletizingVacuumTool against ConveyorBox1, ConveyorBox2, EuroPallet, Half EPAL, LinerStand, StackingTable, near miss 0.05 m
Station logic (signal -> signal, property => property):
  SC_Conveyor1.BoxArrived -> Controler.DI_Box1Arrived
  Controler.DO_Cup21 -> SC_Gripper.Grip
  SC_Conveyor2.BoxArrived -> Controler.DI_Box2Arrived
  SC_Conveyor1.EuroPalletReplacedOut -> Controler.DI_EuroPalletReplaced
  Controler.DO_EuroPalletFull -> SC_Conveyor1.EuroPalletFull
  Controler.DO_HalfPalletFull -> SC_Conveyor2.HalfPalletFull
  SC_Conveyor2.HalfPalletReplacedOut -> Controler.DI_HalfPalletReplaced
  Controler.DO_LinerStackEmpty -> SC_Liners.LinerStackEmpty
  SC_Liners.LinersRefilledOut -> Controler.DI_LinersRefilled
  SC_Conveyor2.HalfPalletReplacedOut -> SC_Liners.PalletReplaced
Targets, tools, work objects and paths stored in the station and not in the controller backup, written as RAPID:
! task T_ROB1
MODULE PalletProgram
  PROC Path_10()
    MoveL PickConveyor2,v1000,z100,toolVacuum\WObj:=wobjConveyor2;
    MoveL PlaceTable,v1000,z100,toolVacuum\WObj:=wobjTable;
    MoveL PickTableStack,v1000,z100,toolVacuum\WObj:=wobjTable;
    MoveL PickLiner,v1000,z100,toolVacuum\WObj:=wobjLinerStack;
    MoveL PlaceHalfPallet,v1000,z100,toolVacuum\WObj:=wobjHalfPallet;
    MoveL PlaceLiner,v1000,z100,toolVacuum\WObj:=wobjHalfPallet;
    MoveL PickConveyor1,v1000,z100,toolVacuum\WObj:=wobjConveyor1;
    MoveL PlaceEuroRow2,v1000,z100,toolVacuum\WObj:=wobjEuroPallet;
    MoveL PlaceEuroRow4,v1000,z100,toolVacuum\WObj:=wobjEuroPallet;
  ENDPROC
ENDMODULE


--- Controller Data/Controler/RAPID/TASK1/PROGMOD/CalibData.mod ---
MODULE CalibData
    !-----------------------------------------------------------------------
	! Tools and work object
	!-----------------------------------------------------------------------
    TASK PERS wobjdata wobjEuroPallet:=[FALSE,TRUE,"",[[600,600,144],[0.707106781,0,0,-0.707106781]],[[0,0,0],[1,0,0,0]]];
    TASK PERS wobjdata wobjHalfPallet:=[FALSE,TRUE,"",[[400,-600,144],[0,0,0,1]],[[0,0,0],[1,0,0,0]]];
    TASK PERS wobjdata wobjConveyor1:=[FALSE,TRUE,"",[[338.5,670,768],[0.707106781,0,0,0.707106781]],[[0,0,0],[1,0,0,0]]];
    TASK PERS wobjdata wobjConveyor2:=[FALSE,TRUE,"",[[-353.5,670,768],[0.707106781,0,0,0.707106781]],[[0,0,0],[1,0,0,0]]];
    TASK PERS wobjdata wobjTable:=[FALSE,TRUE,"",[[-600,600,770],[0,0,0,1]],[[55,170,0],[1,0,0,0]]];
    TASK PERS wobjdata wobjLinerStack:=[FALSE,TRUE,"",[[-500,-160,500],[0,0,0,1]],[[0,0,0],[1,0,0,0]]];
    TASK PERS tooldata toolVacuum:=[TRUE,[[0,0,175],[1,0,0,0]],[1,[0,0,1],[1,0,0,0],0,0,0]];
    ! toolVacuum: mass and CoG are provisional (1 kg), to be estimated

    !-----------------------------------------------------------------------
	! Load data
	!-----------------------------------------------------------------------
    ! Payloads: CoG relative to the TCP of toolVacuum; inertia set to 0 (point mass) until confirmed
    TASK PERS loaddata loadBox1:=[2,[0,0,100],[1,0,0,0],0,0,0];
    ! Box 2 is picked with one corner cup (x=-160, y=-100); on the table fill rows ascending Y, each row descending X
    TASK PERS loaddata loadBox2:=[0.4,[-160,-100,100],[1,0,0,0],0,0,0];
    ! 3x2 stack of box 2 (390 x 260 x 200 mm, 6 x 0.4 kg)
    TASK PERS loaddata loadBox2Stack:=[2.4,[0,0,100],[1,0,0,0],0,0,0];
    ! Liner: corrugated cardboard, 0.8 x 0.54 x 0.01 m3 x 120 kg/m3 = 0.52 kg
    TASK PERS loaddata loadLiner:=[0.52,[0,0,5],[1,0,0,0],0,0,0];
ENDMODULE

--- Controller Data/Controler/RAPID/TASK1/PROGMOD/PalletProgram.mod ---
MODULE PalletProgram

    !***********************************************************************
    ! Industrial Robotics and Offline Programming G1F - University of Skovde
    ! Offline programming project: Pallet Project - Group 2 (JMPM)
    ! Authors: Peru Mendivil and Joaquin Moreno
    ! Robot :   ABB IRB 1600-10/1.45, IRC5 RobotWare 6.13.02 (RobotStudio 2025)
    ! Tool  :   toolVacuum, vacuum gripper with 6 cups (one valve per cup)
    ! Date:    2026-10-30
    !
    ! The robot palletizes two products coming on two conveyors.
    ! Box 1 goes from conveyor 1 to the Euro pallet: 4-2 pattern,
    ! 2 layers (12 boxes). Box 2 goes from conveyor 2 to the stacking
    ! table, where a 3x2 block is formed. The block is then moved to the
    ! half pallet: 2x2 blocks per layer, 3 layers (72 boxes), with a liner
    ! after layers 1 and 2. When both conveyors have a box, the robot
    ! alternates box 1 and box 2. A full pallet is replaced by the operator
    ! from outside the fence, and the robot keeps working with the other
    ! product. With the half pallet full, one block can still be finished
    ! on the table, and it waits there. If the liner stack is empty, the
    ! robot keeps working until a liner is needed; then box 2 waits until
    ! the operator refills the stack.
    !
    ! Structure: Main is a state machine (grafcet). It initialises the
    ! signals and then decides each cycle which box to handle, from the
    ! conveyor sensors, the full-pallet flags and the last box handled.
    ! Each product has its own routine with a finite-state machine for
    ! the place positions. Every place position is calculated with Offs
    ! from one base target per station. ApproachPoint does every
    ! pick/place: approach, vacuum on/off and GripLoad. Work objects,
    ! tool and loads are in the module CalibData.
    !
    ! Naming: VAR, PERS and parameters in camelCase (can change);
    ! CONST, PROC, FUNC and MODULE in PascalCase (fixed).
    !***********************************************************************

    !-----------------------------------------------------------------------
    ! Base targets
    !-----------------------------------------------------------------------
    CONST jointtarget Home:=[[0,0,0,0,90,0],[9E+09,9E+09,9E+09,9E+09,9E+09,9E+09]];

    ! Box 1
    CONST robtarget PickConveyor1:=[[249.5,0,200],[0,0,1,0],[0,0,0,0],[9E+09,9E+09,9E+09,9E+09,9E+09,9E+09]];
    CONST robtarget PlaceEuroRow4:=[[225,525,200],[0,-0.707106781,0.707106781,0],[-2,0,0,0],[9E+09,9E+09,9E+09,9E+09,9E+09,9E+09]];
    CONST robtarget PlaceEuroRow2:=[[350,150,200],[0,1,0,0],[-2,0,-1,0],[9E+09,9E+09,9E+09,9E+09,9E+09,9E+09]];

    ! Box 2
    CONST robtarget PickConveyor2:=[[-35.5,-160,200],[0,-0.707106781,0.707106781,0],[0,0,0,0],[9E+09,9E+09,9E+09,9E+09,9E+09,9E+09]];
    CONST robtarget PlaceTable:=[[-95,165,200],[0,0,1,0],[0,0,0,0],[9E+09,9E+09,9E+09,9E+09,9E+09,9E+09]];
    CONST robtarget PickTableStack:=[[195,130,200],[0,0,1,0],[0,0,0,0],[9E+09,9E+09,9E+09,9E+09,9E+09,9E+09]];
    CONST robtarget PlaceHalfPallet:=[[205,170,200],[0,0,1,0],[0,0,0,0],[9E+09,9E+09,9E+09,9E+09,9E+09,9E+09]];

    ! Liners
    CONST robtarget PickLiner:=[[400,270,100],[0,0,1,0],[0,0,0,0],[9E+09,9E+09,9E+09,9E+09,9E+09,9E+09]];
    CONST robtarget PlaceLiner:=[[400,300,210],[0,0,1,0],[0,0,0,0],[9E+09,9E+09,9E+09,9E+09,9E+09,9E+09]];

    !-----------------------------------------------------------------------
    ! Speeds and heights
    !-----------------------------------------------------------------------
    CONST speeddata TransitSpeed:=v1000;
    CONST speeddata ApproachSpeed:=v300;

    ! Height of every station (world)
    CONST num ConveyorsHeight:=768;
    CONST num TableHeight:=770;
    CONST num LinerStandHeight:=500;
    CONST num EuroPalletHeight:=144;
    CONST num HalfPalletHeight:=144;

    CONST num Box1Height:=200;
    CONST num Box2Height:=200;

    ! Heights for the approach points
    CONST num TransitHeight:=1100;
    CONST num PalletOffsetHeight:=250;
    CONST num MinApproachHeight:=250;

    ! Station identifiers for ApproachHeight
    CONST num StationConveyor1:=1;
    CONST num StationConveyor2:=2;
    CONST num StationTable:=3;
    CONST num StationLinerStand:=4;
    CONST num StationHalfPallet:=5;
    CONST num StationEuroPallet:=6;

    !-----------------------------------------------------------------------
    ! Vacuum gripper
    !-----------------------------------------------------------------------
    CONST num VacuumTime:=1;
    CONST bool CupsAllOn{6}:=[TRUE,TRUE,TRUE,TRUE,TRUE,TRUE];
    CONST bool CupsAllOff{6}:=[FALSE,FALSE,FALSE,FALSE,FALSE,FALSE];
    CONST bool CupsBox2On{6}:=[FALSE,FALSE,FALSE,TRUE,FALSE,FALSE];
    VAR bool cupsState{6}:=[FALSE,FALSE,FALSE,FALSE,FALSE,FALSE];
    VAR signaldo cupSignals{6};

    !-----------------------------------------------------------------------
    ! Box selection
    !-----------------------------------------------------------------------
    CONST num Box1:=1;
    CONST num Box2:=2;
    ! Last box handled, to alternate box 1 and box 2
    VAR num lastBox:=Box2;

    !-----------------------------------------------------------------------
    ! Box 1 state machine parameters and variables
    !-----------------------------------------------------------------------
    CONST num Box1Pos1:=1;
    CONST num Box1Pos2:=2;
    CONST num Box1Pos3:=3;
    CONST num Box1Pos4:=4;
    CONST num Box1Pos5:=5;
    CONST num Box1LastPos:=6;
    CONST num Box1MaxLayers:=2;
    ! Distance between boxes in the row of 4 and in the row of 2
    CONST num EuroRow4Offset:=250;
    CONST num EuroRow2Offset:=500;

    VAR num box1State:=1;
    VAR num box1Layer:=1;
    VAR bool euroPalletFull:=FALSE;

    !-----------------------------------------------------------------------
    ! Box 2 state machine parameters and variables (table)
    !-----------------------------------------------------------------------
    CONST num Box2Pos1:=1;
    CONST num Box2Pos2:=2;
    CONST num Box2Pos3:=3;
    CONST num Box2Pos4:=4;
    CONST num Box2Pos5:=5;
    CONST num Box2LastPos:=6;
    ! Distance between boxes 2 on the table
    CONST num Box2Offset:=130;

    VAR num box2State:=1;
    VAR bool tableFull:=FALSE;

    !-----------------------------------------------------------------------
    ! TransferStack parameters and variables (half pallet)
    !-----------------------------------------------------------------------
    CONST num BlockPos1:=1;
    CONST num BlockPos2:=2;
    CONST num BlockPos3:=3;
    CONST num BlockPos4:=4;
    CONST num Box2MaxLayers:=3;
    ! Distance between 3x2 blocks on the half pallet
    CONST num BlockOffsetX:=3*Box2Offset;
    CONST num BlockOffsetY:=2*Box2Offset;

    VAR num blockState:=1;
    VAR num box2Layer:=1;
    VAR bool halfPalletFull:=FALSE;

    !-----------------------------------------------------------------------
    ! Liners parameters and variables
    !-----------------------------------------------------------------------
    CONST num TotalLiners:=10;
    CONST num LinerHeight:=10;

    VAR num linersLeft:=TotalLiners;
    ! Liner stack empty: warning to the operator, the robot keeps working
    VAR bool linerStackEmpty:=FALSE;
    ! Layer complete but the liner stack is empty: box 2 waits for the refill
    VAR bool linerMissing:=FALSE;

    !-----------------------------------------------------------------------
    ! Main: choose the box and check the operator signals
    !-----------------------------------------------------------------------
    PROC Main()

        InitSignals;
        VacuumControl CupsAllOff;
        SetDO DO_EuroPalletFull,0;
        SetDO DO_HalfPalletFull,0;
        SetDO DO_LinerStackEmpty,0;
        GripLoad load0;
        MoveAbsJ Home,v100,fine,toolVacuum;

        WHILE TRUE DO

            ! Alternate box 1 and box 2 when both are ready
            IF Box1Ready() AND ((NOT Box2Ready()) OR lastBox=Box2) THEN
                ProcessBox1;
            ELSEIF Box2Ready() THEN
                ProcessBox2;
            ENDIF

            ! Half pallet replaced: counters first, then the waiting block
            IF halfPalletFull AND DI_HalfPalletReplaced=1 THEN
                box2Layer:=1;
                blockState:=BlockPos1;
                halfPalletFull:=FALSE;
                SetDO DO_HalfPalletFull,0;
                IF tableFull THEN
                    TransferStack;
                    tableFull:=FALSE;
                ENDIF
            ENDIF

            ! Liner stack refilled: place the missing liner and the waiting block
            IF linerStackEmpty AND DI_LinersRefilled=1 THEN
                linersLeft:=TotalLiners;
                linerStackEmpty:=FALSE;
                SetDO DO_LinerStackEmpty,0;
                IF linerMissing THEN
                    linerMissing:=FALSE;
                    PlaceLayerLiner;
                    IF tableFull THEN
                        TransferStack;
                        tableFull:=FALSE;
                    ENDIF
                ENDIF
            ENDIF

            ! Euro pallet replaced
            IF euroPalletFull AND DI_EuroPalletReplaced=1 THEN
                box1Layer:=1;
                ! Not necessary but safe
                box1State:=Box1Pos1;
                euroPalletFull:=FALSE;
                SetDO DO_EuroPalletFull,0;
            ENDIF
            WaitTime 0.1;
        ENDWHILE
    ENDPROC

    !-----------------------------------------------------------------------
    ! Box ready to be handled
    !-----------------------------------------------------------------------
    FUNC bool Box1Ready()
        ! Box 1 waiting on conveyor 1 and room on the Euro pallet
        RETURN (DI_Box1Arrived=1) AND (NOT euroPalletFull);
    ENDFUNC

    FUNC bool Box2Ready()
        ! Box 2 waiting on conveyor 2 and room on the table
        RETURN (DI_Box2Arrived=1) AND (NOT tableFull);
    ENDFUNC

    !-----------------------------------------------------------------------
    ! Box 1 state machine: conveyor 1 to the Euro pallet
    !-----------------------------------------------------------------------
    PROC ProcessBox1()
        ! Z of the current layer on the Euro pallet
        VAR num layerZ;

        ApproachPoint PickConveyor1,wobjConveyor1,CupsAllOn,loadBox1,ApproachHeight(StationConveyor1);

        layerZ:=(box1Layer-1)*Box1Height;
        TEST box1State
        CASE Box1Pos1:
            ApproachPoint Offs(PlaceEuroRow4,0,0,layerZ),wobjEuroPallet,CupsAllOff,load0,ApproachHeight(StationEuroPallet);
            box1State:=Box1Pos2;
        CASE Box1Pos2:
            ApproachPoint Offs(PlaceEuroRow4,EuroRow4Offset,0,layerZ),wobjEuroPallet,CupsAllOff,load0,ApproachHeight(StationEuroPallet);
            box1State:=Box1Pos3;
        CASE Box1Pos3:
            ApproachPoint Offs(PlaceEuroRow4,2*EuroRow4Offset,0,layerZ),wobjEuroPallet,CupsAllOff,load0,ApproachHeight(StationEuroPallet);
            box1State:=Box1Pos4;
        CASE Box1Pos4:
            ApproachPoint Offs(PlaceEuroRow4,3*EuroRow4Offset,0,layerZ),wobjEuroPallet,CupsAllOff,load0,ApproachHeight(StationEuroPallet);
            box1State:=Box1Pos5;
        CASE Box1Pos5:
            ApproachPoint Offs(PlaceEuroRow2,0,0,layerZ),wobjEuroPallet,CupsAllOff,load0,ApproachHeight(StationEuroPallet);
            box1State:=Box1LastPos;
        CASE Box1LastPos:
            ApproachPoint Offs(PlaceEuroRow2,EuroRow2Offset,0,layerZ),wobjEuroPallet,CupsAllOff,load0,ApproachHeight(StationEuroPallet);
            IF box1Layer=Box1MaxLayers THEN
                euroPalletFull:=TRUE;
                SetDO DO_EuroPalletFull,1;
            ELSE
                Incr box1Layer;
            ENDIF
            box1State:=Box1Pos1;
        DEFAULT:
            box1State:=Box1Pos1;
        ENDTEST
        lastBox:=Box1;
    ENDPROC

    !-----------------------------------------------------------------------
    ! Box 2 state machine: conveyor 2 to the table
    !-----------------------------------------------------------------------
    PROC ProcessBox2()

        ApproachPoint PickConveyor2,wobjConveyor2,CupsBox2On,loadBox2,ApproachHeight(StationConveyor2);

        ! Far row (y=130) first and x from high to low: the box carried never crosses the boxes already placed
        TEST box2State
        CASE Box2Pos1:
            ApproachPoint Offs(PlaceTable,2*Box2Offset,Box2Offset,0),wobjTable,CupsAllOff,load0,ApproachHeight(StationTable);
            box2State:=Box2Pos2;
        CASE Box2Pos2:
            ApproachPoint Offs(PlaceTable,Box2Offset,Box2Offset,0),wobjTable,CupsAllOff,load0,ApproachHeight(StationTable);
            box2State:=Box2Pos3;
        CASE Box2Pos3:
            ApproachPoint Offs(PlaceTable,0,Box2Offset,0),wobjTable,CupsAllOff,load0,ApproachHeight(StationTable);
            box2State:=Box2Pos4;
        CASE Box2Pos4:
            ApproachPoint Offs(PlaceTable,2*Box2Offset,0,0),wobjTable,CupsAllOff,load0,ApproachHeight(StationTable);
            box2State:=Box2Pos5;
        CASE Box2Pos5:
            ApproachPoint Offs(PlaceTable,Box2Offset,0,0),wobjTable,CupsAllOff,load0,ApproachHeight(StationTable);
            box2State:=Box2LastPos;
        CASE Box2LastPos:
            ApproachPoint Offs(PlaceTable,0,0,0),wobjTable,CupsAllOff,load0,ApproachHeight(StationTable);
            IF halfPalletFull OR linerMissing THEN
                tableFull:=TRUE;
            ELSE
                TransferStack;
            ENDIF
            box2State:=Box2Pos1;
        DEFAULT:
            box2State:=Box2Pos1;
        ENDTEST
        lastBox:=Box2;
    ENDPROC

    !-----------------------------------------------------------------------
    ! Box 2: move the 3x2 block from the table to the half pallet
    !-----------------------------------------------------------------------
    PROC TransferStack()
        ! Z of the current layer on the half pallet (block and liner)
        VAR num layerZ;

        ! Pick all 6 boxes 2
        ApproachPoint PickTableStack,wobjTable,CupsAllOn,loadBox2Stack,ApproachHeight(StationTable);

        ! Place group of boxes
        layerZ:=HalfPalletLayerZ();
        TEST blockState
        CASE BlockPos1:
            ApproachPoint Offs(PlaceHalfPallet,0,BlockOffsetY,layerZ),wobjHalfPallet,CupsAllOff,load0,ApproachHeight(StationHalfPallet);
            blockState:=BlockPos2;
        CASE BlockPos2:
            ApproachPoint Offs(PlaceHalfPallet,BlockOffsetX,BlockOffsetY,layerZ),wobjHalfPallet,CupsAllOff,load0,ApproachHeight(StationHalfPallet);
            blockState:=BlockPos3;
        CASE BlockPos3:
            ApproachPoint Offs(PlaceHalfPallet,0,0,layerZ),wobjHalfPallet,CupsAllOff,load0,ApproachHeight(StationHalfPallet);
            blockState:=BlockPos4;
        CASE BlockPos4:
            ApproachPoint Offs(PlaceHalfPallet,BlockOffsetX,0,layerZ),wobjHalfPallet,CupsAllOff,load0,ApproachHeight(StationHalfPallet);
            IF box2Layer=Box2MaxLayers THEN
                halfPalletFull:=TRUE;
                SetDO DO_HalfPalletFull,1;
            ELSEIF linerStackEmpty THEN
                linerMissing:=TRUE;
            ELSE
                PlaceLayerLiner;
            ENDIF
            blockState:=BlockPos1;
        DEFAULT:
            blockState:=BlockPos1;
        ENDTEST
    ENDPROC

    !-----------------------------------------------------------------------
    ! Liner on the layer just finished, then the next layer starts
    !-----------------------------------------------------------------------
    PROC PlaceLayerLiner()
        ApproachPoint Offs(PickLiner,0,0,-(TotalLiners-linersLeft)*LinerHeight),wobjLinerStack,CupsAllOn,loadLiner,ApproachHeight(StationLinerStand);
        ApproachPoint Offs(PlaceLiner,0,0,HalfPalletLayerZ()),wobjHalfPallet,CupsAllOff,load0,ApproachHeight(StationHalfPallet);
        Incr box2Layer;
        Decr linersLeft;
        IF linersLeft=0 THEN
            linerStackEmpty:=TRUE;
            SetDO DO_LinerStackEmpty,1;
        ENDIF
    ENDPROC

    !-----------------------------------------------------------------------
    ! Z of the current layer on the half pallet (block and liner)
    !-----------------------------------------------------------------------
    FUNC num HalfPalletLayerZ()
        ! One liner under every layer except the first one
        RETURN (box2Layer-1)*(Box2Height+LinerHeight);
    ENDFUNC

    !-----------------------------------------------------------------------
    ! Pick or place at a target: approach, vacuum, GripLoad and go up
    !-----------------------------------------------------------------------
    PROC ApproachPoint(robtarget target,PERS wobjdata wobj,bool cups{*},PERS loaddata load,num approachHeight)
        ! cups: cups on/off at the target, load: load after the target
        MoveJ Offs(target,0,0,approachHeight),TransitSpeed,z10,toolVacuum\WObj:=wobj;
        MoveL target,ApproachSpeed,fine,toolVacuum\WObj:=wobj;
        VacuumControl cups;
        GripLoad load;
        MoveL Offs(target,0,0,approachHeight),ApproachSpeed,z10,toolVacuum\WObj:=wobj;
    ENDPROC

    !-----------------------------------------------------------------------
    ! Calculation of approach heights (how much the robot goes up over the target)
    !-----------------------------------------------------------------------
    FUNC num ApproachHeight(num station)
        VAR num approachingHeight:=9E+09;
        TEST station
        CASE StationConveyor1:
            approachingHeight:=TransitHeight-ConveyorsHeight-Box1Height;
        CASE StationConveyor2:
            approachingHeight:=TransitHeight-ConveyorsHeight-Box2Height;
        CASE StationTable:
            approachingHeight:=TransitHeight-TableHeight-Box2Height;
        CASE StationLinerStand:
            approachingHeight:=TransitHeight-LinerStandHeight-linersLeft*LinerHeight;
        CASE StationHalfPallet:
            approachingHeight:=TransitHeight-HalfPalletHeight-HalfPalletLayerZ()-Box2Height-PalletOffsetHeight;
            IF approachingHeight<MinApproachHeight THEN
                approachingHeight:=MinApproachHeight;
            ENDIF
        CASE StationEuroPallet:
            approachingHeight:=TransitHeight-EuroPalletHeight-Box1Height*box1Layer-PalletOffsetHeight;
            IF approachingHeight<MinApproachHeight THEN
                approachingHeight:=MinApproachHeight;
            ENDIF
        DEFAULT:
            ! If another station is entered the robot will announce an error trying to reach 9E+09: Safety stop
        ENDTEST
        RETURN approachingHeight;
    ENDFUNC

    !-----------------------------------------------------------------------
    ! Assignment of logical cup signals with physical signals
    !-----------------------------------------------------------------------
    PROC InitSignals()
        ! Call it first: VacuumControl needs it
        AliasIO DO_Cup11,cupSignals{1};
        AliasIO DO_Cup12,cupSignals{2};
        AliasIO DO_Cup13,cupSignals{3};
        AliasIO DO_Cup21,cupSignals{4};
        AliasIO DO_Cup22,cupSignals{5};
        AliasIO DO_Cup23,cupSignals{6};
    ENDPROC

    !-----------------------------------------------------------------------
    ! Control of the vacuum of every cup
    !-----------------------------------------------------------------------
    PROC VacuumControl(bool cups{*})
        cupsState:=cups;

        FOR i FROM 1 TO Dim(cups,1) DO
            IF cups{i} THEN
                SetDO cupSignals{i},1;
            ELSE
                SetDO cupSignals{i},0;
            ENDIF
        ENDFOR

        ! Robot stopped in position, wait for the vacuum
        WaitTime\InPos,VacuumTime;
    ENDPROC

ENDMODULE

--- Controller Data/Controler/SYSPAR/EIO.cfg ---
EIO:CFG_1.0:6:1::
#
EIO_SIGNAL:

      -Name "DO_Cup11" -SignalType "DO" -Label "Vacuum valve gripper"\
      -Category "Gripper"

      -Name "DI_Box1Arrived" -SignalType "DI" -Label "Box 1 sensor conveyor 1"\
      -Category "Conveyor"

      -Name "DI_Box2Arrived" -SignalType "DI" -Label "Box 2 sensor conveyor 2"\
      -Category "Conveyor"

      -Name "DI_EuroPalletReplaced" -SignalType "DI"\
      -Label "Operator confirms new euro pallet" -Category "Operator"

      -Name "DI_HalfPalletReplaced" -SignalType "DI"\
      -Label "Operator confirms new half pallet" -Category "Operator"

      -Name "AI_VacuumPressure" -SignalType "AI"\
      -Label "Vacuum pressure sensor (bar)" -Category "Gripper" -MaxLog 10

      -Name "DO_Cup12" -SignalType "DO" -Label "Vacuum valve gripper"\
      -Category "Gripper"

      -Name "DO_Cup13" -SignalType "DO" -Label "Vacuum valve gripper"\
      -Category "Gripper"

      -Name "DO_Cup21" -SignalType "DO" -Label "Vacuum valve gripper"\
      -Category "Gripper"

      -Name "DO_Cup22" -SignalType "DO" -Label "Vacuum valve gripper"\
      -Category "Gripper"

      -Name "DO_Cup23" -SignalType "DO" -Label "Vacuum valve gripper"\
      -Category "Gripper"

      -Name "DI_LinersRefilled" -SignalType "DI"\
      -Label "Indicates refilled liners" -Category "Liners"

      -Name "DO_EuroPalletFull" -SignalType "DO"

      -Name "DO_HalfPalletFull" -SignalType "DO"

      -Name "DO_LinerStackEmpty" -SignalType "DO"
